SUBAPPLICATION Uebung_094b5b_AX (* Wie Uebung_094b5_AX, aber mit MyLib::sys::Checkbox_TO_AD2_2 als wiederverwendbarem Baustein statt der einzeln verdrahteten Checkbox_IDA_TO_AX/ASSEMBLE_AD_FROM_AX/AD_TO_AD2/SPLIT_AD_INTO_AX/AX_TO_Checkbox-Kette. *)
  (* Standard: 61499-2; Description: Copyright (c) 2026 Meisterschulen am Ostbahnhof This program and the accompanying materials are made available under the terms of the Eclipse Public License 2.0 which is available at https://www.eclipse.org/legal/epl-2.0/ SPDX-License-Identifier: EPL-2.0 *)
  (* Version 1.0, 2026-10-13, Franz Höpfinger, Meisterschulen am Ostbahnhof, 2. Version von Uebung_094b5_AX: alles ausser AOption_AD_DEMUX_2/OptionalGroup_001/OptionalGroup_002 wurde nach MyLib::sys::Checkbox_TO_AD2_2 ausgelagert. *)
  PACKAGE Uebungen;
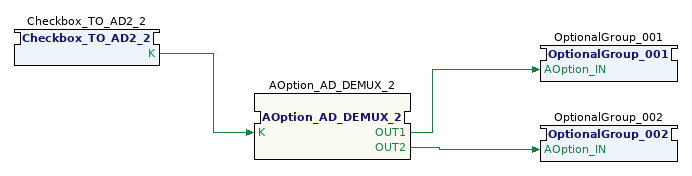
  FBS
    AOption_AD_DEMUX_2 : Option::selection::AOption_AD_DEMUX_2;
  END_FBS
  SUBAPPS
    Checkbox_TO_AD2_2 : MyLib::sys::Checkbox_TO_AD2_2;
    OptionalGroup_001 : MyLib_AX_Option::sys::OptionalGroup_001;
    OptionalGroup_002 : MyLib_AX_Option::sys::OptionalGroup_002;
  END_SUBAPPS
  ADAPTER_CONNECTIONS
    Checkbox_TO_AD2_2.K TO AOption_AD_DEMUX_2.K;
    AOption_AD_DEMUX_2.OUT1 TO OptionalGroup_001.AOption_IN;
    AOption_AD_DEMUX_2.OUT2 TO OptionalGroup_002.AOption_IN;
  END_CONNECTIONS
END_SUBAPPLICATION
